# EPICS autosave request: utcaApp/Db/ebpm_pos_calc.req
$(P)$(R)PosKx-SP
$(P)$(R)PosKy-SP
$(P)$(R)PosKq-SP
$(P)$(R)PosKsum-SP
$(P)$(R)PosXOffset-SP
$(P)$(R)PosYOffset-SP
$(P)$(R)PosQOffset-SP
$(P)$(R)XYPosCal-Sel
$(P)$(R)SumPosCal-Sel
$(P)$(R)QPosCal-Sel
